Fanuc KAREL source: kb00163.compact.KL

PROGRAM KB00163
%STACKSIZE=65535
%PRIORITY=65535
%NOLOCKGROUP
VAR
P1 : FILE
P2 : INTEGER
BEGIN
P2=1
SET_FILE_ATR(P1,P2,1)
END KB00163
